# EPICS autosave request: iocs/meascomp/db/measCompAnalogIn_settings.req
$(P)$(R)Range
$(P)$(R)Type
$(P)$(R)Rate
$(P)$(R).LOPR
$(P)$(R).HOPR
$(P)$(R).EGUF
$(P)$(R).EGUL
$(P)$(R).PREC
$(P)$(R).SCAN
